Staubli VAL3: Lab2A_new.pjx

--- Lab2A_new.pjx ---
parameters version=s6.8 stackSize=5000 millimeterUnit=true
program file=start.pgx
program file=pickAndPlace.pgx
program file=stop.pgx
program file=physicalIO.pgx
data file=Lab2A_new.dtx
alias name=io interface=io autoload=true

--- Lab2A_new.dtx ---


--- start.pgx ---
program start()
// Lab2A Level 3 - shared manual simulation / physical cycle
  local num rowIndex
  local num columnIndex
  local num targetIndex
  local pointRs targetPose
begin
  // ============================================================
  // LAB 2A - NIVEL 3: MISMO CICLO PARA SIMULACION Y FISICO
  // ============================================================
  // ANTES de arrancar: simulation=true manual; false estacion real.
  // Se fija el modo al arrancar: no cambia durante este ciclo.
  // materialType: 0=no metalica roja/derecha; 1=metalica.
  // Matriz VACIA al arrancar: cuatro piezas de cada material.
  userPage()
  cls()
  physicalRun = !simulation

  // ============================================================
  // 2. REINICIAR CONTADORES Y PREPARAR LAS ORDENES
  // ============================================================
  // cycleStep indica en que fase estamos. No lo cambias tu.
  // placedCount[0]: piezas NO metalicas colocadas.
  // placedCount[1]: piezas metalicas colocadas.
  cycleStep = 0
  placedCount[0] = 0
  placedCount[1] = 0

  // Estados iniciales. Barrera retiene las piezas.
  // En simulacion estas son simplemente variables observables.
  // En fisico el adaptador copiara sus valores a las salidas.
  vacuumOn = false
  blowOn = false
  trolleyOn = false
  nonMetalGate = false
  metalGate = false
  barrierClosed = true
  ioReady = false

  // ============================================================
  // 3. CONECTAR LAS VARIABLES CON EL HARDWARE SI ES FISICO
  // ============================================================
  // physicalIO es una tarea que trabaja en paralelo:
  // lee sensores reales y aplica nuestras ordenes a las salidas.
  //
  // Esto permite que los sensores sigan actualizandose mientras
  // el programa principal esta detenido en un wait().
  //
  // En simulacion no creamos esa tarea: los sensores los cambias tu.
  ioReady = false

  if physicalRun
    taskCreate "physicalIO", 10, physicalIO()

    // No continuar hasta que el adaptador haya completado
    // su primera lectura de entradas y escritura de salidas.
    wait(ioReady == true)
    putln("Lab2A_new - PHYSICAL")
  else
    putln("Lab2A_new - MANUAL SIMULATION")
  endIf


  // ============================================================
  // 4. PREPARAR LOS PARAMETROS DE MOVIMIENTO
  // ============================================================
  // moveSpeed agrupa velocidad, aceleracion y deceleracion.
  // blend=off evita redondear las transiciones entre movimientos.
  // Ademas esperaremos a terminar cada movimiento antes de seguir.
  moveSpeed.vel = 10
  moveSpeed.accel = 10
  moveSpeed.decel = 10
  moveSpeed.blend = off


  // ============================================================
  // 5. CALCULAR LA MATRIZ DE DOS FILAS Y CUATRO COLUMNAS
  // ============================================================
  // Referencias ensenadas: placePose[0] para fila 0 y placePose[4] para fila 1.
  // Se conservan ambas joints y se calculan las otras tres columnas por fila.
  //
  // Distribucion de los indices:
  // Primera fila:  0, 1, 2, 3.
  // Segunda fila:  4, 5, 6, 7.
  //
  // Para aplicar distancias en milimetros:
  // 1. Convertimos la joint de referencia a un punto cartesiano.
  // 2. Desplazamos ese punto en Y para recorrer las columnas.
  // 3. Convertimos el resultado de nuevo a joints.

  for rowIndex = 0 to 1
    for columnIndex = 0 to 3
      targetIndex = 4*rowIndex + columnIndex

      // Obtener la posicion del TCP correspondiente a la joint
      // de referencia de SU fila, expresada respecto al sistema world.
      // 4*rowIndex vale 0 para la primera fila y 4 para la segunda.
      targetPose = jointToPoint(vacuumTool, world, placePose[4*rowIndex])

      // Segunda fila: usar su joint ensenada, NO desplazar X=-70.
      // Columnas separadas 60 mm desde la referencia de cada fila.
      // Avance invertido a world Y positiva; verificar destino 1 y 5 en SRS.
      targetPose.trsf.y = targetPose.trsf.y + 60*columnIndex

      // Argumento 1: herramienta cuyo TCP queremos posicionar.
      // Argumento 2: joints de referencia para buscar la solucion.
      // Argumento 3: posicion y orientacion deseadas del TCP.
      // Argumento 4: variable donde se guardan las joints calculadas.
      // Devuelve true si encuentra solucion. No mueve el robot.
      // Columna cero: conservar la joint ensenada (indice 0 o 4).
      // Otras columnas: calcular usando la referencia de su propia fila.
      if columnIndex != 0
        if !pointToJoint(vacuumTool, placePose[4*rowIndex], targetPose, placePose[targetIndex])
          putln("ERROR: unreachable matrix destination")
          putln(targetIndex)
          return
        endIf
      endIf

      // Crear tambien una aproximacion 50 mm por encima del
      // destino. Servira para entrar y salir de forma lineal.
      targetPose.trsf.z = targetPose.trsf.z + 50

      if !pointToJoint(vacuumTool, placePose[targetIndex], targetPose, placeApproach[targetIndex])
        putln("ERROR: unreachable matrix approach")
        putln(targetIndex)
        return
      endIf

    endFor
  endFor

  // ============================================================
  // 6. COLOCAR EL ROBOT EN LA POSICION INICIAL
  // ============================================================
  // movej mueve las articulaciones hasta homePose.
  // El recorrido del TCP no tiene por que ser una linea recta.
  // Esperamos a que termine antes de comenzar la alimentacion.
  movej(homePose, vacuumTool, moveSpeed)
  waitEndMove()


  // ============================================================
  // 7. REPETIR EL CICLO HASTA TENER CUATRO PIEZAS DE CADA TIPO
  // ============================================================
  // materialType=0: NO metalica, roja, rampa derecha.
  // materialType=1: metalica, segunda rampa.
  // El "or" hace que continuemos mientras falte completar
  // cualquiera de los dos materiales.
  // Alimentacion continua durante toda la mision, incluso con el robot ocupado.
  // La barrera dosifica la liberacion; no paramos bOut2 entre piezas.
  trolleyOn = true
  while placedCount[0] < 4 or placedCount[1] < 4

    // ==========================================================
    // FASE 20: LLEVAR LA PIEZA HASTA CLASIFICACION
    // ==========================================================
    // La alimentacion ya esta en marcha. Esperamos presencia bIn1.
    // El material se lee cuando la pieza llega a clasificacion.
    //
    // SIMULACION, en este orden:
    // 1. partIsMetal=false para roja o true para metalica.
    // 2. partAtClass=true: ya esta en clasificacion.
    cycleStep = 20
    putln("20 - Set partIsMetal, then partAtClass=true")
    wait(partAtClass == true)

    // Interpretamos el detector inductivo solo despues de
    // confirmar que hay una pieza delante de el.
    // Guardamos el material para el resto de esta pieza:
    // aunque luego el sensor cambie, materialType ya esta elegido.
    if partIsMetal
      materialType = 1
    else
      materialType = 0
    endIf

    // Aunque su fila ya este llena, dejamos pasar esta pieza.
    // La decision de recoger se toma despues, usando el mismo contador.

    // ==========================================================
    // FASE 30: ORDENAR LA RUTA Y DAR TIEMPO AL ACTUADOR
    // ==========================================================
    // Estas dos variables son ORDENES:
    // nonMetalGate controla bOut3, actuador 1.
    // metalGate controla bOut4, actuador 2.
    //
    // La comparacion produce true o false directamente:
    // - No metalica: nonMetalGate=true, metalGate=false.
    // - Metalica: nonMetalGate=false, metalGate=true.
    //
    // TODO FISICO: confirmar que salida=1 significa empujar
    // y que estas combinaciones conducen a la rampa correcta.
    cycleStep = 30
    putln("30 - Select route; actuator settling delay")

    nonMetalGate = materialType == 0
    metalGate = materialType == 1

    // Suponemos que los actuadores alcanzan su posicion.
    // No leemos ni esperamos finales de carrera bIn5..bIn8.
    // Dejamos una pausa antes de liberar la pieza.
    // TODO FISICO: ajustar 0.5 s al tiempo real de los actuadores.
    // Esta pausa NO confirma que el actuador se haya movido.
    delay(0.5)

    // ==========================================================
    // FASE 40: ABRIR BREVEMENTE Y CERRAR ANTES DE ESPERAR LA RAMPA
    // ==========================================================
    // La cinta sigue en marcha. No podemos dejar la barrera abierta
    // hasta que la pieza llegue a bIn4: pasarian tambien las demas.
    // Damos un pulso de apertura y ordenamos cerrar inmediatamente.
    // Retener=true envia bOut5=0; liberar=false envia bOut5=1.
    // TODO FISICO: verificar polaridad y pulso de 0.4 s para UNA pieza.
    // El pulso es temporal: por si solo no confirma dosificacion unitaria.
    cycleStep = 40
    putln("40 - Barrier pulse; then wait partAtRamp=true")


    barrierClosed = false
    delay(0.4)
    barrierClosed = true

    // delay para copiar la order al pin
    delay(0.05)
    if barrierClosed
      putln("40 - after cllose: barrierClosed=true")
    else
      putln("40 - after cllose: barrierClosed=false")
    endIf
    if io:bOut5
      putln("40 - after cllose: bOut5=true")
    else
      putln("40 - after cllose: bOut5=false")
    endIf

    // La barrera ya tiene orden de cierre durante esta espera.
    // SIMULACION: partAtRamp=true representa el paso de la pieza.
    wait(partAtRamp == true)

    // ==========================================================
    // FASE 50: ESPERAR QUE LA PIEZA DEJE LIBRE EL SENSOR DE RAMPA
    // ==========================================================
    // No esperamos partAtClass=false: con la cinta continua,
    // la siguiente pieza puede estar ya retenida en clasificacion.
    // Su material se leera en la siguiente vuelta, no en esta.
    cycleStep = 50
    putln("50 - Wait: partAtRamp=false")
    wait(partAtRamp == false)

    // El detector confirma PASO, no llegada al punto de recogida.
    // En fisico dejamos un tiempo adicional para que llegue.
    if physicalRun
      delay(0.5)
    endIf


    // ==========================================================
    // RECOGER SOLO SI QUEDAN HUECOS PARA ESTE MATERIAL
    // ==========================================================
    // La pieza ya ha pasado por su rampa. Si su fila esta completa,
    // no movemos el robot, no calculamos otro indice y no contamos.
    // Volvemos a clasificar la siguiente hasta completar ambas filas.
    if placedCount[materialType] < 4
      // No metalicas: destinos 0..3. Metalicas: destinos 4..7.
      placeIndex = 4*materialType + placedCount[materialType]
      call pickAndPlace()
      placedCount[materialType] = placedCount[materialType] + 1
      cycleStep = 80
      putln("80 - Piece placed; next classification part")
    else
      cycleStep = 80
      putln("80 - Row full: part passed without pickup; next part")
    endIf
  endWhile

  // ============================================================
  // MISION COMPLETADA
  // ============================================================
  // Llegamos aqui cuando ambos contadores valen cuatro.
  trolleyOn = false
  barrierClosed = true
  cycleStep = 100
  putln("100 - Completed: four parts of each material")
end

--- physicalIO.pgx ---
program physicalIO()
// Lab2A Level 3 - shared manual simulation / physical cycle
begin
  // ============================================================
  // ADAPTADOR ENTRE LAS VARIABLES Y LOS PINES FISICOS
  // ============================================================
  // start solo crea esta tarea cuando simulation=false.
  //
  // Trabaja en paralelo con el ciclo principal:
  // 1. Lee entradas reales y actualiza nuestros sensores bool.
  // 2. Lee nuestras ordenes bool y las escribe en salidas reales.
  // 3. Hace una pausa breve y repite.
  //
  // Asi, un wait del programa principal puede desbloquearse
  // cuando esta tarea detecta un cambio en un sensor real.
  //
  // En fisico NO modificar los sensores bool a mano:
  // esta tarea los sobrescribe con las lecturas reales.
  while true
    // ==========================================================
    // 1. LEER LOS SENSORES DE PIEZA
    // ==========================================================
    // Cada comparacion convierte la lectura de la entrada
    // en un valor bool: true si esta activa, false si no.

    // bIn0: confirma que hay una pieza en la ventosa.
    // No es la orden de aspiracion, sino su confirmacion.
    partOnTool = io:bIn0 == true

    // bIn1: confirma presencia en la zona de clasificacion.
    partAtClass = io:bIn1 == true

    // bIn2: detector inductivo.
    // Activo significa metalica.
    // Inactivo se interpreta como no metalica SOLO cuando
    // sabemos que hay una pieza en clasificacion.
    partIsMetal = io:bIn2 == true

    // bIn3 no se usa: esperamos directamente presencia en clasificacion.

    // bIn4: detecta el paso de una pieza por la rampa.
    // No confirma que ya haya llegado al punto de recogida.
    partAtRamp = io:bIn4 == true


    // bIn5..bIn8 no se usan en esta version simplificada.
    // Los desviadores reciben su orden y damos un tiempo fijo.

    // ==========================================================
    // 3. APLICAR LAS ORDENES DE LA VENTOSA
    // ==========================================================
    // El programa principal cambia vacuumOn y blowOn.
    // Aqui convertimos esas variables en salidas fisicas.

    // bOut0: activar o desactivar la aspiracion.
    io:bOut0 = vacuumOn

    // bOut1: activar o desactivar el soplado.
    io:bOut1 = blowOn


    // ==========================================================
    // 4. APLICAR LAS ORDENES DE ALIMENTACION Y CLASIFICACION
    // ==========================================================

    // bOut2: orden al carro de alimentacion.
    io:bOut2 = trolleyOn

    // bOut3: actuador 1, asociado a las no metalicas.
    // TODO FISICO: confirmar que true significa empujar.
    io:bOut3 = nonMetalGate

    // bOut4: actuador 2, asociado a las metalicas.
    // TODO FISICO: confirmar que true significa empujar.
    io:bOut4 = metalGate

    // bOut5: barrera de retencion.
    // Polaridad invertida: retener=true envia bOut5=0.
    // Liberar=false envia bOut5=1; pendiente comprobar en fisico.
    io:bOut5 = !barrierClosed


    // ==========================================================
    // 5. AVISAR DE QUE LA PRIMERA ACTUALIZACION ESTA HECHA
    // ==========================================================
    // start espera esta variable antes de continuar en fisico.
    // Una vez pasa a true, permanece true durante la ejecucion.
    ioReady = true

    // Pausa de 0.01 segundos antes de repetir las lecturas.
    // No garantiza un periodo exacto de 10 ms: tambien cuenta
    // el tiempo empleado en ejecutar y planificar la tarea.
    delay(0.01)

  endWhile
end

--- pickAndPlace.pgx ---
program pickAndPlace()
// Lab2A Level 3 - shared manual simulation / physical cycle
begin
  // ============================================================
  // RECOGER: materialType ELIGE RAMPA; placeIndex ELIGE DESTINO
  // ============================================================
  vacuumOn = false
  blowOn = false
  movej(pickApproach[materialType], vacuumTool, moveSpeed)
  waitEndMove()
  movel(jointToPoint(vacuumTool, world, pickPose[materialType]), vacuumTool, moveSpeed)
  waitEndMove()
  vacuumOn = true
  cycleStep = 60
  putln("60 - Wait: partOnTool=true; keep true during transfer")
  wait(partOnTool == true)
  movel(jointToPoint(vacuumTool, world, pickApproach[materialType]), vacuumTool, moveSpeed)
  waitEndMove()

  // ============================================================
  // TRASLADAR, DEPOSITAR Y CONFIRMAR LIBERACION
  // ============================================================
  movej(placeApproach[placeIndex], vacuumTool, moveSpeed)
  waitEndMove()
  movel(jointToPoint(vacuumTool, world, placePose[placeIndex]), vacuumTool, moveSpeed)
  waitEndMove()
  vacuumOn = false
  blowOn = true
  // TODO FISICO: validar duracion del soplado.
  delay(0.3)
  blowOn = false
  cycleStep = 70
  putln("70 - Wait: partOnTool=false")
  wait(partOnTool == false)

  // ============================================================
  // RETIRAR Y VOLVER A HOME ANTES DE CONTAR LA PIEZA
  // ============================================================
  movel(jointToPoint(vacuumTool, world, placeApproach[placeIndex]), vacuumTool, moveSpeed)
  waitEndMove()
  movej(homePose, vacuumTool, moveSpeed)
  waitEndMove()
end

--- stop.pgx ---
program stop()
// Lab2A Level 3 - shared manual simulation / physical cycle
begin
  // ============================================================
  // 1. REINICIAR EL CONTROL DE MOVIMIENTO
  // ============================================================
  resetMotion()

  // ============================================================
  // 2. PREPARAR LAS ORDENES DE PARADA
  // ============================================================
  // Parar el carro, ordenar que la barrera retenga
  // y dejar de soplar.
  trolleyOn = false
  barrierClosed = true
  blowOn = false

  // ============================================================
  // 3. SI ES FISICO, PARAR EL ADAPTADOR Y ESCRIBIR LAS SALIDAS
  // ============================================================
  if physicalRun
    taskKill("physicalIO")

    // Parar carro y soplado.
    io:bOut2 = false
    io:bOut1 = false

    // Retencion con la nueva polaridad: bOut5=0.
    // Debe coincidir con !barrierClosed del adaptador.
    io:bOut5 = false

    // No escribimos bOut0: conservamos la aspiracion.
    // Tampoco cambiamos aqui los actuadores de clasificacion.
  endIf


  // ============================================================
  // 4. INDICAR QUE SE HA EJECUTADO LA PARADA
  // ============================================================
  cycleStep = -1
  putln("Stopped - empty matrix before a new start")

end
